(* IEC 61131-3 sources: Caravan/Archiv/12-04-19/Stations/MachineControl/MachineControl/Class/HmiStateBit35, 1 file *)

(* ---- HmiStateBit35.st ---- *)
#include "..\..\Source\Common\hmi_nuc.h"

(*!
<Class
	Name               = "HmiStateBit35"
	Revision           = "0.4"
	RealtimeTask       = "false"
	CyclicTask         = "false"
	BackgroundTask     = "false"
	Sigmatek           = "true"
	OSInterface        = "false"
	HighPriority       = "false"
	Automatic          = "false"
	UpdateMode         = "Prescan"
	SharedCommandTable = "true"
	Objectsize         = "(284,120)">
	<Channels>
		<Server Name="ClassSvr" Visualized="false" Initialize="false" WriteProtected="true" Retentive="false"/>
		<Client Name="ChkBit" Required="true" Internal="false"/>
		<Client Name="ComPort" Required="true" Internal="false"/>
		<Client Name="StringLib" Required="true" Internal="false"/>
		<Client Name="VarList" Required="true" Internal="false"/>
	</Channels>
	<Dependencies>
		<Files>
			<File Path=".\Source\Common\hmi_nuc.h" Include="true"/>
		</Files>
	</Dependencies>
	<RevDoku>
		<Owner Company="sigmatek" Author="kolott"/>
		<Dokumentation Revision="0.4" Date="2016-06-28" Author="kolott" Company="sigmatek" Description="Type of membervariable PHmi changen foom ^void to ^LseEasy."/>
		<Dokumentation Revision="0.3" Date="2016-03-07" Author="kolott" Company="sigmatek" Description="unused local variable deleted"/>
		<Dokumentation Revision="0.2" Date="2016-02-04" Author="kolott" Company="sigmatek" Description="new method GetMapCrc() added"/>
		<Dokumentation Revision="0.1" Date="2014-11-26" Author="kolott" Company="sigmatek" Description="EasyMap.xml: enable &apos;_&apos; in statebitname"/>
	</RevDoku>
</Class>
*)
HmiStateBit35 : CLASS
	TYPE
#pragma pack(push, 1)
	  StateBit : STRUCT
	    CBit : HMI_CHKBIT;
	    Value : DINT;
	    Access : UINT;
	  END_STRUCT;
#pragma pack(pop)
	END_TYPE
  //Servers:
	ClassSvr 	: SvrChCmd_DINT;
  //Clients:
	ChkBit 	: CltChCmd_HmiChkBitList;
	ComPort 	: CltChCmd_HmiComPort;
	VarList 	: CltChCmd_HmiVarList;
	StringLib 	: CltChCmd_HmiStrLib;
  //Variables:
		UsedNo 	: UDINT;
		UsedChkBit : ARRAY [0..255] OF StateBit;

		RunIdx 	: UDINT;
		PHmi 	: ^LseEasy;
  //Functions:

	FUNCTION GLOBAL RefreshAll;

	FUNCTION GLOBAL RefreshRun;

	FUNCTION GLOBAL AddEntry
		VAR_INPUT
			pcb 	: ^HMI_CHKBIT;
			access 	: UINT;
			pany 	: ^HMI_ANYTHING;
		END_VAR
		VAR_OUTPUT
			retcode 	: USINT;
		END_VAR;

	FUNCTION GLOBAL Start
		VAR_INPUT
			pthis 	: ^LseEasy;
		END_VAR;

	FUNCTION Seek
		VAR_INPUT
			pcb 	: ^HMI_CHKBIT;
			access 	: UINT;
		END_VAR
		VAR_OUTPUT
			retcode 	: UDINT;
		END_VAR;

	FUNCTION CallEntry
		VAR_INPUT
			idx 	: UDINT;
			update 	: BOOL;
		END_VAR;

	FUNCTION GLOBAL GetVarInfo
		VAR_INPUT
			pany 	: ^HMI_ANYTHING;
		END_VAR
		VAR_OUTPUT
			retcode 	: ^HMI_VARINFO;
		END_VAR;

	FUNCTION GLOBAL GetMapInfoXML
		VAR_INPUT
			index 	: UDINT;
			ptext 	: ^CHAR;
		END_VAR
		VAR_OUTPUT
			retcode 	: ^CHAR;
		END_VAR;

	FUNCTION GLOBAL GetMapCrc
		VAR_OUTPUT
			retcode 	: UDINT;
		END_VAR;
  //Tables:
	FUNCTION @STD
		VAR_OUTPUT
			ret_code	: CONFSTATES;
		END_VAR;
	FUNCTION GLOBAL TAB @CT_;
END_CLASS;

#pragma usingLtd HmiChkBitList
#pragma usingLtd HmiComPort
#pragma usingLtd HmiStrLib
#pragma usingLtd HmiVarList

#pragma usingLtd LseEasy

#includeC "..\LseEasy\Create.h"
#pragma using LseEasy

FUNCTION GLOBAL HmiStateBit35::Start
	VAR_INPUT
		pthis 	: ^LseEasy;
	END_VAR

  PHmi     := pthis;
  UsedNo   := 0;
  RunIdx   := 0;
  ClassSvr := 0;

END_FUNCTION

FUNCTION HmiStateBit35::CallEntry
  VAR_INPUT
  	idx : udint;
  	update : bool;
  END_VAR
  VAR
  	st : dint;
    ph : ^StateBit;
  END_VAR

  if(idx < UsedNo) then

    ph := #UsedChkBit[idx];
    st := 16#FF;

    if(ChkBit.Get(#ph^.CBit) <> nil) then
      if(ChkBit.Call(#ph^.CBit) = false) then
        st := st xor SBIT_VISIBLE;
      end_if;
    end_if;

    if(ph^.Access <> 0) then
      if(PHmi <> NIL) then
        if(PHmi^.HmiAccess(ph^.Access) = false) then
          st := st xor SBIT_ACCESS;
        end_if;
      end_if;
    end_if;

    if((ph^.Value <> st) | (update = true)) then
      if(ComPort.SendStateBit(idx$uint + 1, st$usint) = true) then
        ph^.Value := st;
      end_if;
    end_if;
  end_if;

END_FUNCTION

FUNCTION GLOBAL HmiStateBit35::RefreshAll
  VAR
  	idx : udint;
  END_VAR

  idx := 0;
  while(idx < UsedNo) do
    CallEntry(idx, true);
    idx += 1;
  end_while;

END_FUNCTION

FUNCTION GLOBAL HmiStateBit35::RefreshRun

  if(UsedNo) then
    if(RunIdx >= UsedNo) then
      RunIdx := 0;
    end_if;

    CallEntry(RunIdx, false);

    RunIdx += 1;
  end_if;

END_FUNCTION

FUNCTION HmiStateBit35::Seek
	VAR_INPUT
		pcb 	: ^HMI_CHKBIT;
		access 	: UINT;
	END_VAR
	VAR_OUTPUT
		retcode 	: UDINT;
	END_VAR
  VAR
  	idx : udint;
    ph : ^StateBit;
  END_VAR

  ph  := #UsedChkBit[0];
  idx := 0;
  while(idx < UsedNo) do
    if((ph^.CBit.no = pcb^.no) & (ph^.CBit.invert = pcb^.invert) & (ph^.Access = access)) then
      retcode := idx;
      return;
    end_if;
    ph  += sizeof(StateBit);
    idx += 1;
  end_while;

  retcode := 16#FFFFFFFF;

END_FUNCTION

FUNCTION GLOBAL HmiStateBit35::GetVarInfo
	VAR_INPUT
		pany 	: ^HMI_ANYTHING;
	END_VAR
	VAR_OUTPUT
		retcode 	: ^HMI_VARINFO;
	END_VAR

  retcode := nil;
  if(pany <> nil) then
    if((pany^.ima = HMI_IMA_V_SERVERLIST) | (pany^.ima = HMI_IMA_V_SERVERTEXT00) | (pany^.ima = HMI_IMA_V_SERVERUNITTEXT)) then
      retcode := VarList.Get(pany^.value$udint);
    end_if;
  end_if;

END_FUNCTION

FUNCTION GLOBAL HmiStateBit35::AddEntry
	VAR_INPUT
		pcb 	: ^HMI_CHKBIT;
		access 	: UINT;
		pany 	: ^HMI_ANYTHING;
	END_VAR
	VAR_OUTPUT
		retcode 	: USINT;
	END_VAR
  VAR
  	idx : udint;
    st : bool;
    cbit : HMI_CHKBIT;
    pvi : ^HMI_VARINFO;
  END_VAR

  retcode := 0;
  st      := false;

  if(ChkBit.Get(pcb) <> nil) then
    st := true;
  else
    pvi := GetVarInfo(pany);
    if(pvi <> nil) then
      if(ChkBit.Get(#pvi^.chkbit) <> nil) then
        st  := true;
        pcb := #pvi^.chkbit;
      end_if;
    end_if;

    if(st = false) then
      pcb := #cbit;
      init_HMI_CHKBIT(pcb);
    end_if;
  end_if;

  if(access <> 0) then
    st := true;
  else
    pvi := GetVarInfo(pany);
    if(pvi <> nil) then
      if(pvi^.access <> 0) then
        access := pvi^.access;
        st     := true;
      end_if;
    end_if;
  end_if;

  if(st = true) then
    idx := Seek(pcb, access);
    if(idx > UsedNo) then
      if(UsedNo >= 255) then
        return;
      end_if;

      UsedChkBit[UsedNo].CBit   := pcb^;
      UsedChkBit[UsedNo].Value  := -2244766;
      UsedChkBit[UsedNo].Access := access;
      retcode                   := UsedNo$usint;
      UsedNo                    += 1;
      ClassSvr                  += 1;
    else
      retcode := idx$usint;
    end_if;

    retcode += 1;
  end_if;

END_FUNCTION

FUNCTION GLOBAL HmiStateBit35::GetMapInfoXML
	VAR_INPUT
		index 	: UDINT;
		ptext 	: ^CHAR;
	END_VAR
	VAR_OUTPUT
		retcode 	: ^CHAR;
	END_VAR
  VAR
    psb : ^StateBit;
    ph, plabel : ^char;
  END_VAR

  retcode := nil;
  ph      := ptext;
  if(index < UsedNo) then
    psb := #UsedChkBit[index];

    StringLib.StrCpy(ph, 1, "<statebit id=?", 1);
    ph += StringLib.StrLen(ph, 1);
    StringLib.DintToStr(ph, to_dint(index+1), 16#800, 1);
    StringLib.StrCat(ph, 1, "? sequence=?", 1);
    ph += StringLib.StrLen(ph, 1);

    plabel := ChkBit.GetLabel(#psb^.CBit);
    if(plabel <> nil) then
      if(psb^.CBit.invert) then
        ph^ := '!'; ph  += 1;
      end_if;
      StringLib.StrCpy(ph, 1, plabel, 1);
      ph += StringLib.StrLen(ph, 1);
    end_if;

    if(psb^.Access <> 0) then
      if(plabel <> nil) then
        StringLib.StrCat(ph, 1, " or ", 1);
        ph += StringLib.StrLen(ph, 1);
      end_if;

      StringLib.StrCpy(ph, 1, "(Access", 1);
      ph += StringLib.StrLen(ph, 1);
      StringLib.DintToStr(ph, psb^.Access, 16#800, 1);
      StringLib.StrCat(ph, 1, " shl 1)", 1);
    end_if;

    StringLib.StrCat(ph, 1, "?/>", 1);
    StringLib.StrXchg(ptext, '?', '"');

    retcode := ptext;
  end_if;

END_FUNCTION

FUNCTION GLOBAL HmiStateBit35::GetMapCrc
	VAR_OUTPUT
		retcode 	: UDINT;
	END_VAR
  VAR
  	index, len : udint;
    psb : ^StateBit;
    plabel : ^char;
  END_VAR

  retcode := 0;
  index   := 0;
  while(index < UsedNo) do
    psb   := #UsedChkBit[index];
    index += 1;

    retcode := (retcode rol 1) xor index;

    plabel := ChkBit.GetLabel(#psb^.CBit);
    if(plabel <> nil) then
      len := StringLib.StrLen(plabel, 1) + 1;
      retcode := make_crc32(retcode, plabel, len);
    end_if;

    if(psb^.CBit.invert) then
      retcode := (retcode rol 1) xor 1;
    end_if;

    if(psb^.Access <> 0) then
      retcode := (retcode rol 1) xor psb^.Access;
    end_if;
  end_while;

END_FUNCTION
